(* IEC 61131-3 sources: moqui-plc/simatic-ax/src/moqui/framework/src/main/org/moqui/motion (part 3) *)

                        hasPending := FALSE;
                    END_IF;

                    commandAborted := TRUE;
                    internalStatus := AxisInternalStatus#Ready;
                ELSE
                    pendingCmd := cmd;
                    pendingOldPosition := position; pendingOldDistance := distance; pendingOldVelocity := velocity;
                    pendingOldRatioNumerator := ratioNumerator; pendingOldRatioDenominator := ratioDenominator;
                    pendingOldCamVersion := camVersion; pendingOldStartMode := startMode;
                    pendingOldMasterOffset := masterOffset; pendingOldSlaveOffset := slaveOffset;
                    hasPending := TRUE;
                    oldCmd := pendingCmd;

                    CASE pendingCmd OF
                        AxisCmd#MoveVelocity : moveVelocityExecute := TRUE;
                        AxisCmd#MoveAbsolute : moveAbsoluteExecute := TRUE;
                        AxisCmd#MoveRelative : moveRelativeExecute := TRUE;
                        AxisCmd#MoveAdditive : moveAdditiveExecute := TRUE;
                        AxisCmd#MoveSuperimposed : moveSuperimposedExecute := TRUE;
                        AxisCmd#Halt : haltExecute := TRUE;
                        AxisCmd#GearIn : gearInExecute := TRUE;
                        AxisCmd#GearInPos : gearInPosExecute := TRUE;
                        AxisCmd#CamIn : camInExecute := TRUE;
                        AxisCmd#Phasing : phasingExecute := TRUE;
                        AxisCmd#SetPosition : setPositionExecute := TRUE;
                        AxisCmd#PositionProfile : posProfileExecute := TRUE;
                        AxisCmd#VelocityProfile : velProfileExecute := TRUE;
                        AxisCmd#AccelerationProfile: accProfileExecute := TRUE;
                    ELSE
						hasPending := FALSE;
						commandAborted := TRUE;
						internalStatus := AxisInternalStatus#Ready;
                    END_CASE;
                END_IF;
            END_IF;

        (* ReadParameter *)
        AxisInternalStatus#ReadParameterState :
            IF readParameter.Valid THEN
                readParameterExecute := FALSE;
                parameterReadValue := readParameter.Value;
                commandExecuted := TRUE;
                internalStatus := AxisInternalStatus#Ready;
            END_IF;
            IF cmd <> oldCmd THEN
                readParameterExecute := FALSE;
                commandAborted := TRUE;
                internalStatus := AxisInternalStatus#Ready;
            END_IF;

        (* WriteParameter *)
        AxisInternalStatus#WriteParameterState :
            IF writeParameter.Done THEN
                writeParameterExecute := FALSE;
                commandExecuted := TRUE;
                internalStatus := AxisInternalStatus#Ready;
            END_IF;
            IF cmd <> oldCmd THEN
                writeParameterExecute := FALSE;
                commandAborted := TRUE;
                internalStatus := AxisInternalStatus#Ready;
            END_IF;

        (* ReadBoolParameter *)
        AxisInternalStatus#ReadBoolParameterState :
            IF readBoolParameter.Valid THEN
                readBoolParameterExecute := FALSE;
                parameterBoolRead := readBoolParameter.Value;
                commandExecuted := TRUE;
                internalStatus := AxisInternalStatus#Ready;
            END_IF;
            IF cmd <> oldCmd THEN
                readBoolParameterExecute := FALSE;
                commandAborted := TRUE;
                internalStatus := AxisInternalStatus#Ready;
            END_IF;

        (* WriteBoolParameter *)
        AxisInternalStatus#WriteBoolParameterState :
            IF writeBoolParameter.Done THEN
                writeBoolParameterExecute := FALSE;
                commandExecuted := TRUE;
                internalStatus := AxisInternalStatus#Ready;
            END_IF;
            IF cmd <> oldCmd THEN
                writeBoolParameterExecute := FALSE;
                commandAborted := TRUE;
                internalStatus := AxisInternalStatus#Ready;
            END_IF;

        (* TouchProbe - capture axis position on hardware trigger *)
        AxisInternalStatus#TouchProbeState :
            IF touchProbe.Done THEN
                touchProbeExecute := FALSE;
                touchProbeValue := touchProbe.RecordedPosition;
                commandExecuted := TRUE;
                internalStatus := AxisInternalStatus#Ready;
            END_IF;
            IF cmd <> oldCmd THEN
                touchProbeExecute := FALSE;
                commandAborted := TRUE;
                internalStatus := AxisInternalStatus#Ready;
            END_IF;

        (* AbortTrigger - cancel any pending touch probe *)
        AxisInternalStatus#AbortTriggerState :
            IF abortTrigger.Done THEN
                abortTriggerExecute := FALSE;
                commandExecuted := TRUE;
                internalStatus := AxisInternalStatus#Ready;
            END_IF;
            IF cmd <> oldCmd THEN
                abortTriggerExecute := FALSE;
                commandAborted := TRUE;
                internalStatus := AxisInternalStatus#Ready;
            END_IF;
    END_CASE;

END_IF; (* End error-recovery guard *)

(*
 * Status Handler - level-triggered, unconditional, every cycle
 *)
readActualPosition(
    Axis := slave,
    Enable := TRUE
);
actualPosition := readActualPosition.Position;

readActualVelocity(
    Axis := slave,
    Enable := TRUE
);
actualVelocity := readActualVelocity.Velocity;

readActualTorque(
    Axis := slave,
    Enable := TRUE
);
actualTorque := readActualTorque.Torque;

readAxisError(
    Axis := slave,
    Enable := TRUE
);
axisErrorId := readAxisError.AxisErrorID;

readStatus(
    Axis := slave,
    Enable := TRUE
);
(* Priority order matches PLCopen FSM: ErrorStop > Disabled > Stopping > Homing > motion states > Standstill *)
IF readStatus.ErrorStop THEN
    status := AxisStatus#ErrorStop;
ELSIF readStatus.Disabled THEN
    status := AxisStatus#Disabled;
ELSIF readStatus.Stopping THEN
    status := AxisStatus#Stopping;
ELSIF readStatus.Homing THEN
    status := AxisStatus#Homing;
ELSIF readStatus.SynchronizedMotion THEN
    status := AxisStatus#SynchronizedMotion;
ELSIF readStatus.ContinuousMotion THEN
    status := AxisStatus#ContinuousMotion;
ELSIF readStatus.DiscreteMotion THEN
    status := AxisStatus#DiscreteMotion;
ELSIF readStatus.Standstill THEN
    status := AxisStatus#Standstill;
ELSE
    status := AxisStatus#Standstill; (* Fallback - consider adding Unknown to AxisStatus DUT *)
END_IF;

(*
 * PLCopen FB calls - unconditional every PLC cycle.
 * Execute / Enable signals are generated exclusively by the FSM above.
 * All motion parameters come directly from VAR_INPUT each cycle.
 *)

(* Administrative / Configuration *)
power(
    Axis := slave,
    Enable := powerEnable,
    bRegulatorOn := powerEnable,
    bDriveStart := powerEnable
);

resetCmd(
    Axis := slave,
    Execute := resetCmdExecute
);

setPosition(
    Axis := slave,
    Execute := setPositionExecute,
    Position := position,
    Mode := setPositionMode
);

(* Homing *)
home(
    Axis := slave,
    Execute := homeExecute,
    Position := homePosition
);

(* Motion *)
moveVelocity(
    Axis := slave,
    Execute := moveVelocityExecute,
    Velocity := velocity,
    Acceleration := acceleration,
    Deceleration := deceleration,
    Jerk := jerk,
    Direction := direction,
    BufferMode := bufferMode
);

moveAbsolute(
    Axis := slave,
    Execute := moveAbsoluteExecute,
    Position := position,
    Velocity := velocity,
    Acceleration := acceleration,
    Deceleration := deceleration,
    Jerk := jerk,
    Direction := direction,
    BufferMode := bufferMode
);

moveRelative(
    Axis := slave,
    Execute := moveRelativeExecute,
    Distance := distance,
    Velocity := velocity,
    Acceleration := acceleration,
    Deceleration := deceleration,
    Jerk := jerk,
    BufferMode := bufferMode
);

moveAdditive(
    Axis := slave,
    Execute := moveAdditiveExecute,
    Distance := distance,
    Velocity := velocity,
    Acceleration := acceleration,
    Deceleration := deceleration,
    Jerk := jerk
);

moveSuperimposed(
    Axis := slave,
    Execute := moveSuperimposedExecute,
    Distance := distance,
    VelocityDiff := velocityDiff,
    Acceleration := acceleration,
    Deceleration := deceleration,
    Jerk := jerk
);

halt(
    Axis := slave,
    Execute := haltExecute,
    Deceleration := deceleration,
    Jerk := jerk
);

haltSuperimposed(
    Axis := slave,
    Execute := haltSuperimposedExecute,
    Deceleration := deceleration,
    Jerk := jerk
);

stop(
    Axis := slave,
    Execute := stopExecute,
    Deceleration := deceleration,
    Jerk := jerk
);

jog(
    Axis := slave,
    JogForward := jogForward AND (internalStatus = AxisInternalStatus#JogState),
    JogBackward := jogBackward AND (internalStatus = AxisInternalStatus#JogState),
    Velocity := velocity,
    Acceleration := acceleration,
    Deceleration := deceleration,
    Jerk := jerk
);

(* Override *)
setOverride(
    Axis := slave,
    Enable := overrideEnable,
    VelFactor := velFactor,
    AccFactor := accFactor,
    JerkFactor := jerkFactor
);

(* Synchronization - master reference required *)
IF master <> NULL THEN
    gearIn(
        Master := master,
        Slave := slave,
        Execute := gearInExecute,
        RatioNumerator := ratioNumerator,
        RatioDenominator := TO_UDINT(ratioDenominator),
        Acceleration := acceleration,
        Deceleration := deceleration,
        Jerk := jerk,
        BufferMode := bufferMode
    );
    gearInPos(
        Master := master,
        Slave := slave,
        Execute := gearInPosExecute,
        RatioNumerator := ratioNumerator,
        RatioDenominator := ratioDenominator,
        MasterSyncPosition := masterSyncPos,
        SlaveSyncPosition := slaveSyncPos
    );
    camIn(
        Master := master,
        Slave := slave,
        Execute := camInExecute,
        CamTableID := camId,
        StartMode := startMode,
        MasterOffset := masterOffset,
        SlaveOffset := slaveOffset,
        BufferMode := bufferMode
    );
    phasing(
        Master := master,
        Slave := slave,
        Execute := phasingExecute,
        PhaseShift := phaseShift,
        Velocity := velocity,
        Acceleration := acceleration,
        Deceleration := deceleration,
        Jerk := jerk
    );
END_IF;

gearOut(
    Slave := slave,
    Execute := gearOutExecute
);

camOut(
    Slave := slave,
    Execute := camOutExecute
);

(* Profiles *)
IF positionProfile <> NULL THEN
    mcPositionProfile(
        Axis := slave,
        Execute := posProfileExecute,
        TimePosition := positionProfile
    );
END_IF;

IF velocityProfile <> NULL THEN
    mcVelocityProfile(
        Axis := slave,
        Execute := velProfileExecute,
        TimeVelocity := velocityProfile
    );
END_IF;

IF accelerationProfile <> NULL THEN
    mcAccProfile(
        Axis := slave,
        Execute := accProfileExecute,
        TimeAcceleration := accelerationProfile
    );
END_IF;

(* Parameter access *)
readParameter(
    Axis := slave,
    Enable := readParameterExecute,
    ParameterNumber := parameterNumber
);

writeParameter(
    Axis := slave,
    Execute := writeParameterExecute,
    ParameterNumber := parameterNumber,
    Value := parameterValue
);

readBoolParameter(
    Axis := slave,
    Enable := readBoolParameterExecute,
    ParameterNumber := parameterNumber
);

writeBoolParameter(
    Axis := slave,
    Execute := writeBoolParameterExecute,
    ParameterNumber := parameterNumber,
    Value := parameterBoolValue
);

(* Additional services - triggerInput reference required *)
IF triggerInput <> NULL THEN
    touchProbe(
        Axis := slave,
        Execute := touchProbeExecute,
        TriggerInput := triggerInput,
        WindowOnly := touchProbeWindow,
        FirstPosition := touchProbeFirst,
        LastPosition := touchProbeLast
    );
    abortTrigger(
        Axis := slave,
        Execute := abortTriggerExecute,
        TriggerInput := triggerInput
    );
END_IF;
END_FUNCTION_BLOCK
